(*
SPDX-FileCopyrightText: © 2026 Oleksandr Tiutyk <trofimich@gmail.com>
SPDX-License-Identifier: MIT
License: https://opensource.org/license/mit
*)

(*!
<summary>
Beckhoff counter output control channel process image.
</summary>
<description>
Encapsulates 16-bit control word and 32-bit unsigned preset counter value (SetCounterValue : UDINT) for fast
counter terminals.
When used for I/O, link located fields or their containing buffers to the matching selected PDOs.
The record is not a packed wire buffer; compiler padding is not part of the device specification.
Unlinked/default values do not prove valid I/O. The caller evaluates bus/channel validity before use.
Use one owner task per instance and externally synchronize other access; multi-field snapshots are not atomic.
Copies store data without creating hardware links. Keep borrowed field references valid while consumers are bound.
This passive record performs no validation, synchronization, configuration or protocol advancement.
</description>
*)
TYPE COUNTER_OUTPUT_CHANNEL :
STRUCT
	Control AT %Q* : WORD;
	SetCounterValue AT %Q* : UDINT;
END_STRUCT
END_TYPE

(* stored: Version 1.1.0.1, ProductVersion 3.1.4026.20
   DUT COUNTER_OUTPUT_CHANNEL: Id {59851d15-ecdf-40bd-9291-1262bcc613ff} *)
